FUNCTION_BLOCK FB_StartupControl_Tests EXTENDS TcUnit.FB_TestSuite

Repeated_Request_Is_Dropped_When_Online();
First_Request_Is_Kept();
Init_Gate();
Suspend_Is_Never_Online();
Suspend_Reports_Parked_And_Error();
Conditional_Aborts();
Events_Last_One_Scan();
External_Abort_Input();
Publish_On_Change_And_Heartbeat();
Power_Dropped_Without_Abort_Stays_Initializing();
Stop_On_Accepted_Request_Before_Initializing();

METHOD PRIVATE Repeated_Request_Is_Dropped_When_Online
VAR
    ctl : BROTLib.FB_StartupControl;
    rs : LREAL;
    keep : BOOL;
    ok : BOOL;
END_VAR
TEST('Repeated_Request_Is_Dropped_When_Online');
keep := ctl.BeginScan(Power := TRUE, Ready := FALSE);
ctl.MarkCalibrating();
ctl.MarkCompleted();
rs := ctl.Update(Error := FALSE, Parked := FALSE, Parking := FALSE, Operational := TRUE, AbortExtra := FALSE);
AssertEquals_LREAL(1.0, rs, 0.0001, 'online after completion');
keep := ctl.BeginScan(Power := TRUE, Ready := TRUE);
AssertFalse(keep, 'repeated power request dropped');
rs := ctl.Update(Error := FALSE, Parked := FALSE, Parking := FALSE, Operational := TRUE, AbortExtra := FALSE);
AssertEquals_LREAL(1.0, rs, 0.0001, 'repeat does not restart calibration');
TEST_FINISHED();
END_METHOD

METHOD PRIVATE First_Request_Is_Kept
VAR
    ctl : BROTLib.FB_StartupControl;
    rs : LREAL;
    keep : BOOL;
    ok : BOOL;
END_VAR
TEST('First_Request_Is_Kept');
keep := ctl.BeginScan(Power := TRUE, Ready := FALSE);
AssertTrue(keep, 'first request kept');
rs := ctl.Update(Error := FALSE, Parked := FALSE, Parking := FALSE, Operational := TRUE, AbortExtra := FALSE);
AssertEquals_LREAL(0.7, rs, 0.0001, 'preparation');
AssertTrue(ctl.Initializing, 'initializing output');
TEST_FINISHED();
END_METHOD

METHOD PRIVATE Init_Gate
VAR
    ctl : BROTLib.FB_StartupControl;
    rs : LREAL;
    keep : BOOL;
    ok : BOOL;
END_VAR
TEST('Init_Gate');
AssertTrue(ctl.AcceptInit(), 'idle telescope accepts Init');
keep := ctl.BeginScan(Power := TRUE, Ready := FALSE);
rs := ctl.Update(Error := FALSE, Parked := FALSE, Parking := FALSE, Operational := TRUE, AbortExtra := FALSE);
AssertFalse(ctl.AcceptInit(), 'running startup is joined, not restarted');
ctl.MarkCompleted();
rs := ctl.Update(Error := FALSE, Parked := FALSE, Parking := FALSE, Operational := TRUE, AbortExtra := FALSE);
AssertFalse(ctl.AcceptInit(), 'online telescope ignores Init');
keep := ctl.BeginScan(Power := FALSE, Ready := TRUE);
rs := ctl.Update(Error := FALSE, Parked := FALSE, Parking := FALSE, Operational := FALSE, AbortExtra := FALSE);
AssertEquals_LREAL(-2.0, rs, 0.0001, 'interlock');
AssertFalse(ctl.AcceptInit(), 'Init during an interlock must not recalibrate');
keep := ctl.BeginScan(Power := FALSE, Ready := TRUE);
rs := ctl.Update(Error := FALSE, Parked := FALSE, Parking := FALSE, Operational := TRUE, AbortExtra := FALSE);
AssertEquals_LREAL(1.0, rs, 0.0001, 'recovers without a new startup');
ctl.MarkAborted();
rs := ctl.Update(Error := FALSE, Parked := FALSE, Parking := FALSE, Operational := TRUE, AbortExtra := FALSE);
AssertTrue(ctl.AcceptInit(), 'aborted startup may be requested again');
TEST_FINISHED();
END_METHOD

METHOD PRIVATE Suspend_Is_Never_Online
VAR
    ctl : BROTLib.FB_StartupControl;
    rs : LREAL;
    keep : BOOL;
    ok : BOOL;
END_VAR
TEST('Suspend_Is_Never_Online');
keep := ctl.BeginScan(Power := TRUE, Ready := FALSE);
ctl.MarkCalibrating();
ctl.MarkCompleted();
rs := ctl.Update(Error := FALSE, Parked := FALSE, Parking := FALSE, Operational := TRUE, AbortExtra := FALSE);
AssertEquals_LREAL(1.0, rs, 0.0001, 'online after completion');
ok := ctl.EnterSuspend();
AssertTrue(ok, 'first scan of the suspension');
ok := ctl.EnterSuspend();
AssertFalse(ok, 'only once');
rs := ctl.Suspend(Error := FALSE, Parked := FALSE);
AssertEquals_LREAL(-2.0, rs, 0.0001, 'suspended is not online');
AssertFalse(ctl.AcceptInit(), 'no Init while suspended');
keep := ctl.BeginScan(Power := FALSE, Ready := TRUE);
rs := ctl.Update(Error := FALSE, Parked := FALSE, Parking := FALSE, Operational := TRUE, AbortExtra := FALSE);
AssertEquals_LREAL(-2.0, rs, 0.0001, 'back in automatic mode still needs a new init');
AssertTrue(ctl.AcceptInit(), 'Init accepted again');
TEST_FINISHED();
END_METHOD

METHOD PRIVATE Suspend_Reports_Parked_And_Error
VAR
    ctl : BROTLib.FB_StartupControl;
    rs : LREAL;
    keep : BOOL;
    ok : BOOL;
END_VAR
TEST('Suspend_Reports_Parked_And_Error');
rs := ctl.Suspend(Error := FALSE, Parked := TRUE);
AssertEquals_LREAL(0.0, rs, 0.0001, 'parked');
rs := ctl.Suspend(Error := TRUE, Parked := TRUE);
AssertEquals_LREAL(-1.0, rs, 0.0001, 'error');
TEST_FINISHED();
END_METHOD

METHOD PRIVATE Conditional_Aborts
VAR
    ctl : BROTLib.FB_StartupControl;
    rs : LREAL;
    keep : BOOL;
    ok : BOOL;
END_VAR
TEST('Conditional_Aborts');
keep := ctl.BeginScan(Power := TRUE, Ready := FALSE);
ctl.MarkCalibrating();
ctl.MarkCompleted();
rs := ctl.Update(Error := FALSE, Parked := FALSE, Parking := FALSE, Operational := TRUE, AbortExtra := FALSE);
AssertEquals_LREAL(1.0, rs, 0.0001, 'online after completion');
ctl.MarkAbortedIfInitializing();
ctl.MarkAbortedIfStarting(Power := FALSE);
rs := ctl.Update(Error := FALSE, Parked := FALSE, Parking := FALSE, Operational := TRUE, AbortExtra := FALSE);
AssertEquals_LREAL(1.0, rs, 0.0001, 'a stop on an online telescope is not a startup abort');
ctl.MarkAbortedIfStarting(Power := TRUE);
rs := ctl.Update(Error := FALSE, Parked := FALSE, Parking := FALSE, Operational := TRUE, AbortExtra := FALSE);
AssertEquals_LREAL(-2.0, rs, 0.0001, 'pending power request aborted');
keep := ctl.BeginScan(Power := TRUE, Ready := FALSE);
rs := ctl.Update(Error := FALSE, Parked := FALSE, Parking := FALSE, Operational := TRUE, AbortExtra := FALSE);
ctl.MarkAbortedIfInitializing();
rs := ctl.Update(Error := FALSE, Parked := FALSE, Parking := FALSE, Operational := TRUE, AbortExtra := FALSE);
AssertEquals_LREAL(-2.0, rs, 0.0001, 'running startup aborted');
TEST_FINISHED();
END_METHOD

METHOD PRIVATE Events_Last_One_Scan
VAR
    ctl : BROTLib.FB_StartupControl;
    rs : LREAL;
    keep : BOOL;
    ok : BOOL;
END_VAR
TEST('Events_Last_One_Scan');
keep := ctl.BeginScan(Power := TRUE, Ready := FALSE);
ctl.MarkAborted();
rs := ctl.Update(Error := FALSE, Parked := FALSE, Parking := FALSE, Operational := TRUE, AbortExtra := FALSE);
AssertEquals_LREAL(-2.0, rs, 0.0001, 'abort wins');
keep := ctl.BeginScan(Power := TRUE, Ready := FALSE);
rs := ctl.Update(Error := FALSE, Parked := FALSE, Parking := FALSE, Operational := TRUE, AbortExtra := FALSE);
AssertEquals_LREAL(0.7, rs, 0.0001, 'abort of the previous scan is gone');
TEST_FINISHED();
END_METHOD

METHOD PRIVATE External_Abort_Input
VAR
    ctl : BROTLib.FB_StartupControl;
    rs : LREAL;
    keep : BOOL;
    ok : BOOL;
END_VAR
TEST('External_Abort_Input');
keep := ctl.BeginScan(Power := TRUE, Ready := FALSE);
ctl.MarkCalibrating();
ctl.MarkCompleted();
rs := ctl.Update(Error := FALSE, Parked := FALSE, Parking := FALSE, Operational := TRUE, AbortExtra := FALSE);
AssertEquals_LREAL(1.0, rs, 0.0001, 'online after completion');
rs := ctl.Update(Error := FALSE, Parked := FALSE, Parking := FALSE, Operational := TRUE, AbortExtra := TRUE);
AssertEquals_LREAL(-2.0, rs, 0.0001, 'E-stop style abort');
TEST_FINISHED();
END_METHOD

METHOD PRIVATE Publish_On_Change_And_Heartbeat
VAR
    ctl : BROTLib.FB_StartupControl;
    rs : LREAL;
    keep : BOOL;
    ok : BOOL;
END_VAR
TEST('Publish_On_Change_And_Heartbeat');
rs := ctl.Update(Error := FALSE, Parked := TRUE, Parking := FALSE, Operational := FALSE, AbortExtra := FALSE);
AssertFalse(ctl.PublishDue(CommValid := FALSE, Heartbeat := FALSE), 'no comm, nothing sent');
AssertTrue(ctl.PublishDue(CommValid := TRUE, Heartbeat := FALSE), 'first value, and the missed one is still due');
AssertFalse(ctl.PublishDue(CommValid := TRUE, Heartbeat := FALSE), 'unchanged');
AssertTrue(ctl.PublishDue(CommValid := TRUE, Heartbeat := TRUE), 'heartbeat repeats the value');
keep := ctl.BeginScan(Power := TRUE, Ready := FALSE);
rs := ctl.Update(Error := FALSE, Parked := FALSE, Parking := FALSE, Operational := TRUE, AbortExtra := FALSE);
AssertTrue(ctl.PublishDue(CommValid := TRUE, Heartbeat := FALSE), 'change');
TEST_FINISHED();
END_METHOD

METHOD PRIVATE Power_Dropped_Without_Abort_Stays_Initializing
VAR
    ctl : BROTLib.FB_StartupControl;
    rs : LREAL;
    keep : BOOL;
END_VAR
TEST('Power_Dropped_Without_Abort_Stays_Initializing');
// MONETcommon #80: bPower dropped by an error without an abort leaves the startup stuck until stop/reset
keep := ctl.BeginScan(Power := TRUE, Ready := FALSE);
ctl.MarkCalibrating();
rs := ctl.Update(Error := FALSE, Parked := FALSE, Parking := FALSE, Operational := TRUE, AbortExtra := FALSE);
AssertEquals_LREAL(0.8, rs, 0.0001, 'calibrating');
keep := ctl.BeginScan(Power := FALSE, Ready := FALSE);
rs := ctl.Update(Error := FALSE, Parked := FALSE, Parking := FALSE, Operational := TRUE, AbortExtra := FALSE);
AssertEquals_LREAL(0.8, rs, 0.0001, 'dropped power alone does not leave the startup');
AssertFalse(ctl.AcceptInit(), 'a new power-on is refused while stuck');
ctl.MarkAbortedIfStarting(Power := FALSE);
rs := ctl.Update(Error := FALSE, Parked := FALSE, Parking := FALSE, Operational := TRUE, AbortExtra := FALSE);
AssertEquals_LREAL(-2.0, rs, 0.0001, 'stop aborts the stuck startup');
AssertFalse(ctl.Initializing, 'no longer initializing');
AssertTrue(ctl.AcceptInit(), 'power-on accepted again');
TEST_FINISHED();
END_METHOD

METHOD PRIVATE Stop_On_Accepted_Request_Before_Initializing
VAR
    ctl : BROTLib.FB_StartupControl;
    rs : LREAL;
    keep : BOOL;
END_VAR
TEST('Stop_On_Accepted_Request_Before_Initializing');
keep := ctl.BeginScan(Power := TRUE, Ready := FALSE);
ctl.MarkAbortedIfStarting(Power := TRUE);
rs := ctl.Update(Error := FALSE, Parked := FALSE, Parking := FALSE, Operational := TRUE, AbortExtra := FALSE);
AssertEquals_LREAL(-2.0, rs, 0.0001, 'stop wins over a request accepted in the same scan');
AssertFalse(ctl.Initializing, 'never initializing');
TEST_FINISHED();
END_METHOD

END_FUNCTION_BLOCK

(* stored: Version 1.1.0.1, ProductVersion 3.1.4024.15
   POU FB_StartupControl_Tests: Id {cceb447c-dfa7-4da9-9aa4-bb8b76cf91d5}, SpecialFunc None
   Method Repeated_Request_Is_Dropped_When_Online: Id {f55a2374-8991-498c-9e2a-386f87d993e6}
   Method First_Request_Is_Kept: Id {1f7bafa1-3fc1-4a17-a502-68814f9386f3}
   Method Init_Gate: Id {6716ed97-a58c-4f52-a528-7b5de711dd8e}
   Method Suspend_Is_Never_Online: Id {c7683e92-4400-45b6-8d02-f6c15a5421d4}
   Method Suspend_Reports_Parked_And_Error: Id {956dd5a9-042d-41e2-91bd-15f9f79d7f38}
   Method Conditional_Aborts: Id {9b65ae49-20f4-44ea-b5a6-216332b3d7e8}
   Method Events_Last_One_Scan: Id {82931cb8-60d9-4ce7-9ce9-147a86575277}
   Method External_Abort_Input: Id {6276b5d2-b16c-4d23-9bd1-6c383d0e0277}
   Method Publish_On_Change_And_Heartbeat: Id {85f10240-ac7a-40de-b1d4-68dae42023d9}
   Method Power_Dropped_Without_Abort_Stays_Initializing: Id {f5016899-1182-4cc1-a807-e194aee85fb3}
   Method Stop_On_Accepted_Request_Before_Initializing: Id {b3e945c0-dbfb-4768-b228-135e7c8e643e} *)
